Fanuc KAREL source: KT00743.KL

PROGRAM KT00743
%NOLOCKGROUP
VAR
  ARG: ARRAY[4] OF VECTOR
  OUT: INTEGER
BEGIN
  OUT = ARRAY_LEN(ARG)
END KT00743
